Fanuc KAREL source: kd00068.KL

-- PROVISIONAL review KL for V770-1; original PC SHA256 97f14b5dfe7aa7ed92f710c1da10f49a582991522895c8e2eb04d2fbef89891e
-- Incomplete behavior may be omitted. Consult companion uncertainty JSON. Do not deploy.
PROGRAM KD00068
%NOLOCKGROUP
VAR
  I : INTEGER
  J : INTEGER
  B : BOOLEAN
  R : REAL
  S : STRING[80]
BEGIN
  -- UNRESOLVED_PC offsets 5-29; opcodes 9D,81,18,9D,1B,9D,12,2E,1B,2E,13,04
  -- UNRESOLVED_PC offsets 34-38; opcodes 7F
END KD00068
